(* IEC 61131-3 sources: codesys-framework/txt/application/WeVe Core (library)/80 Command/FB_Command, 9 files *)

(* ---- Abort.method.st ---- *)
// Het actieve commando afbreken (Stop, QuickStop, mode-wissel).
METHOD Abort
VAR_INPUT
END_VAR

// --- BEGIN IMPLEMENTATION ---

IF _eResult = E_CommandResult.Busy THEN
	_eResult := E_CommandResult.Aborted;
END_IF

(* ---- Active.prop.st ---- *)
PROPERTY Active : INT
// --- BEGIN IMPLEMENTATION ---

// ----------- GET -----------
VAR
END_VAR

// -- BEGIN IMPLEMENTATION GET --
IF _eResult = E_CommandResult.Busy THEN
	Active := _iActive;
ELSE
	Active := 0;
END_IF

(* ---- Cyclic.method.st ---- *)
// 1x per cyclus aanroepen in de body van de module, vóór de uitvoering.
// Bij een timeout wordt het commando hier al Error, zodat de uitvoering in dezelfde cyclus stopt.
METHOD Cyclic
VAR_INPUT
END_VAR

// --- BEGIN IMPLEMENTATION ---

_xPolledPrev := _xPolled;
_xPolled := FALSE;

// Timeout: timer loopt enkel zolang het commando Busy is en er een timeout is ingesteld
_fbTimeout(IN := _eResult = E_CommandResult.Busy AND _tTimeout > T#0S, PT := _tTimeout);

IF _fbTimeout.Q THEN
	_eResult := E_CommandResult.Error;
	_xTimedOut := TRUE;
END_IF

(* ---- Fail.method.st ---- *)
// Door de module: het actieve commando is gefaald. De module meldt zelf de oorzaak.
METHOD Fail
VAR_INPUT
END_VAR

// --- BEGIN IMPLEMENTATION ---

IF _eResult = E_CommandResult.Busy THEN
	_eResult := E_CommandResult.Error;
END_IF

(* ---- Finish.method.st ---- *)
// Door de module: het actieve commando is goed afgewerkt.
METHOD Finish
VAR_INPUT
END_VAR

// --- BEGIN IMPLEMENTATION ---

IF _eResult = E_CommandResult.Busy THEN
	_eResult := E_CommandResult.Done;
END_IF

(* ---- Invoke.method.st ---- *)
// Start een commando, of geeft de status terug als het al loopt.
// xStart is 1 cyclus TRUE wanneer het commando effectief start: neem dan de parameters over.
//
// Een eindresultaat (Done, Error, Aborted) wordt maar 1x afgeleverd aan wie doorlopend pollt.
// De volgende Invoke van hetzelfde commando start het dus opnieuw, ook in de onmiddellijk
// volgende stap (bv. twee keer Move na elkaar met een andere positie).
// Daarom: maximaal 1x per cyclus aanroepen, en verder gaan zodra er een eindresultaat is.
METHOD Invoke : E_CommandResult
VAR_INPUT
	iCmd 		: INT;		// commando-id uit de enum van de module, > 0 (0 = geen commando)
	xAllowed 	: BOOL;		// mag de module nu starten? (bv. enabled, geen fout)
	tTimeout 	: TIME := T#0S;		// max duur van het commando, T#0S = geen timeout
END_VAR
VAR_OUTPUT
	xStart 		: BOOL;
END_VAR
// --- BEGIN IMPLEMENTATION ---

_xPolled := TRUE;

// Ongeldig commando-id: weigeren, nooit stil negeren
IF iCmd <= 0 THEN
	Invoke := E_CommandResult.Rejected;
	RETURN;
END_IF

IF iCmd = _iActive THEN

	// Loopt nog: pollen
	IF _eResult = E_CommandResult.Busy THEN
		Invoke := E_CommandResult.Busy;
		RETURN;
	END_IF

	// Eindresultaat, vorige cyclus nog gepold en nog niet afgeleverd: 1x afleveren
	IF _xPolledPrev AND NOT _xDelivered THEN
		_xDelivered := TRUE;
		Invoke := _eResult;
		RETURN;
	END_IF

END_IF

// Ander commando bezig of module niet klaar: weigeren, nooit stil negeren
IF _eResult = E_CommandResult.Busy OR NOT xAllowed THEN
	Invoke := E_CommandResult.Rejected;
	RETURN;
END_IF

// Starten
_iActive := iCmd;
_eResult := E_CommandResult.Busy;
_xDelivered := FALSE;
_tTimeout := tTimeout;
_xTimedOut := FALSE;
_fbTimeout(IN := FALSE);	// timer van het vorige commando resetten
xStart := TRUE;
Invoke := E_CommandResult.Busy;

(* ---- Last.prop.st ---- *)
// Laatst gestarte commando, ook als het al klaar, gefaald of verlopen is. 0 = nog nooit iets gestart.
PROPERTY Last : INT
// --- BEGIN IMPLEMENTATION ---

// ----------- GET -----------
VAR
END_VAR

// -- BEGIN IMPLEMENTATION GET --
Last := _iActive;

(* ---- ResultOf.method.st ---- *)
// Resultaat van een commando opvragen zonder iets te starten.
// Blijft staan tot er een nieuw commando start. Idle = dit commando is niet het laatste.
METHOD ResultOf : E_CommandResult
VAR_INPUT
	iCmd 	: INT;
END_VAR
// --- BEGIN IMPLEMENTATION ---

IF iCmd = _iActive THEN
	ResultOf := _eResult;
ELSE
	ResultOf := E_CommandResult.Idle;
END_IF

(* ---- TimedOut.prop.st ---- *)
// TRUE als het laatste commando gefaald is door de timeout. Blijft staan tot er een nieuw commando start.
// Bedoeld voor een event in de module: _fbEvents.Condition(..., xCondition := _fbCmd.TimedOut, ...).
PROPERTY TimedOut : BOOL
// --- BEGIN IMPLEMENTATION ---

// ----------- GET -----------
VAR
END_VAR

// -- BEGIN IMPLEMENTATION GET --
TimedOut := _xTimedOut;
